// TIA Portal V21 export
// export: Created 2026-11-07T17:04:59.5495749Z, ExportSetting WithDefaults, DisplayName Totally Integrated Automation Portal, DisplayVersion V21, DisplayName STEP 7 Professional, DisplayVersion V21, DisplayName STEP 7 Safety, DisplayVersion V21, DisplayName Tech WebApplication, DisplayVersion V21, DisplayName WinCC Basic/Comfort/Advanced, DisplayVersion V21, DisplayName WinCC Unified, DisplayVersion V21
TextList "TL_State"  ListRange=Decimal
  TextListEntry   EntryType=SingleValue, Text="ISKLJUČENO"
  TextListEntry   EntryType=SingleValue, From=1, To=1, Text="INICIJALIZACIJA"
  TextListEntry   EntryType=SingleValue, From=2, To=2, Text="SPREMAN"
  TextListEntry   EntryType=SingleValue, From=3, To=3, Text="RADI"
  TextListEntry   EntryType=SingleValue, From=4, To=4, Text="PAUZA"
  TextListEntry   EntryType=SingleValue, From=5, To=5, Text="ALARM"
  TextListEntry   EntryType=SingleValue, From=6, To=6, Text="ZAVRŠENO"
  TextListEntry   EntryType=SingleValue, From=7, To=7, Text="PLANIRANJE"
